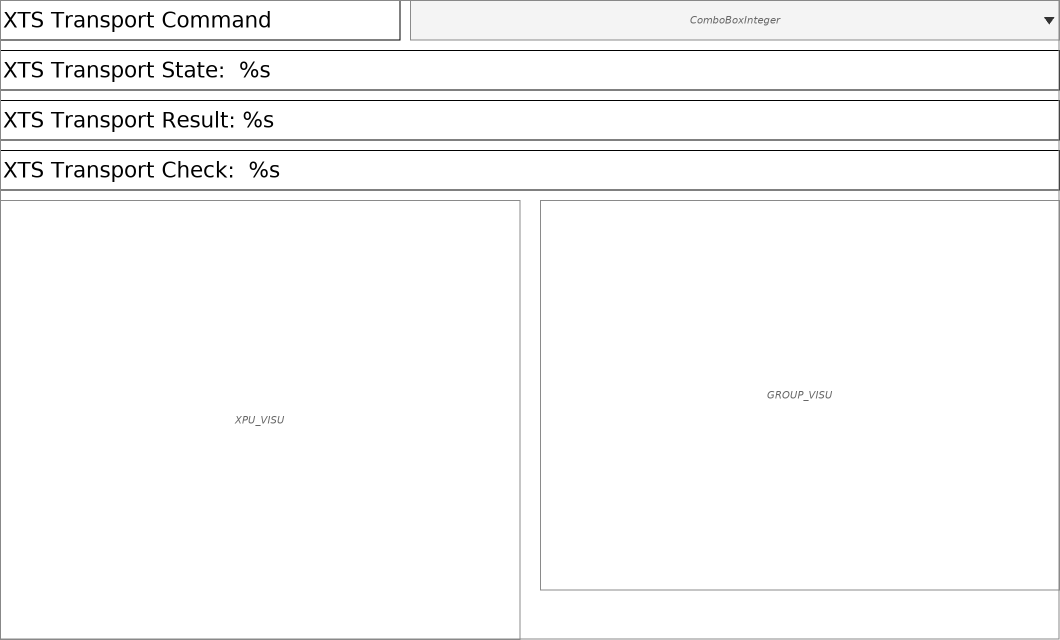
VISUALIZATION TRANSPORT_VISU  // 1060x640
VAR_IN_OUT
	Data    : ST_VISU_POOL;
END_VAR
    Rectangle (0,0 400x40), "XTS Transport Command"
    ComboBoxInteger (410,0 650x40), variable: GVL_XTS.XtsTransportCtrl.Cmd, text list: 'TL_E_CTRL_TRANSPORT'
    Rectangle (0,50 1060x40), "XTS Transport State: %s", text variable: Data.sTransportState
    Rectangle (0,100 1060x40), "XTS Transport Result: %s", text variable: Data.sTransportResult
    Rectangle (0,150 1060x40), "XTS Transport Check: %s", text variable: Data.sTransportCheck
    Frame (0,200 520x440)
        shows XPU_VISU(stXpuState := GVL_XTS.XtsTransportState.XpuState, stXpuInfo := GVL_XTS.XtsTransportState.XpuInfo, stXpuStrings := Data.stXpuStrings)
    Frame (540,200 520x390)
        shows GROUP_VISU(stGroupInfo := GVL_XTS.XtsTransportState.GroupInfo, sGroupState := Data.sCaGroupState)
END_VISUALIZATION

(* stored: Version 1.1.0.1, ProductVersion 3.1.4026.20
   Visu TRANSPORT_VISU: Id {f55b8ab6-35e1-44dc-8419-64447d714789} *)
